ABB RobotStudio station: TPL2_Heredia_Biancuzzo.rspag

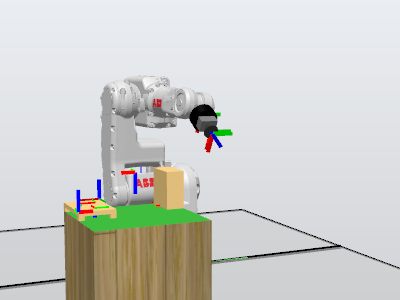
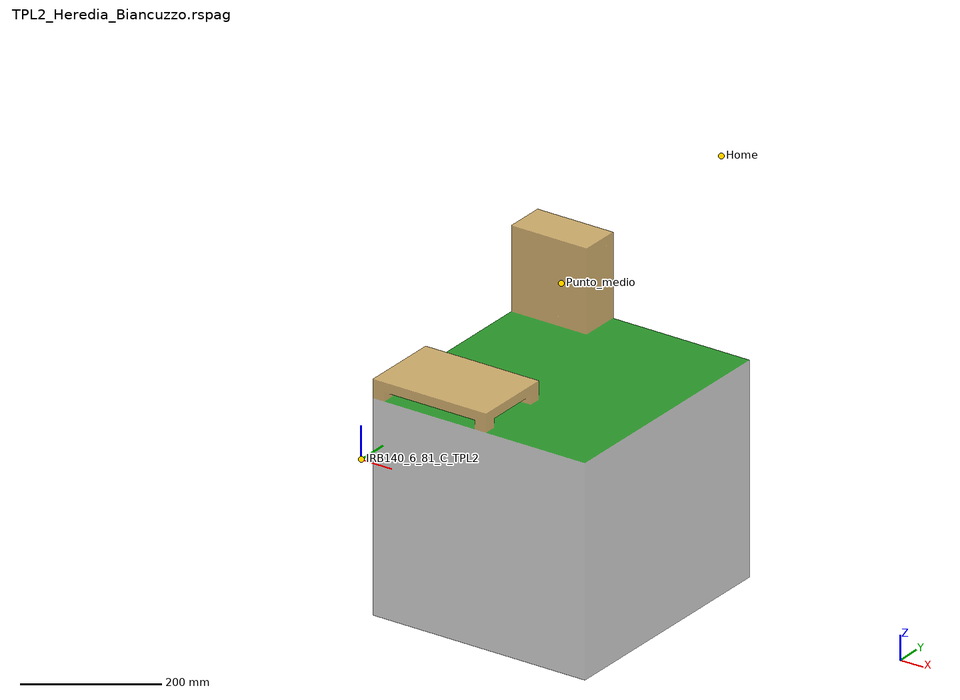
[picture v1: parts stored in the station drawn from their meshes, with robot base, taught points and paths (robot models come from the ABB library and are not in the file)]
--- station ---
Station Paletizado (saved by RobotStudio 25.5.11605.0)
Controller IRB140_6_81_TPL2
  mechanical unit ROB_1: IRB140_6_81_C_TPL2, 6 joints, base frame (0, 0, 0) mm
Layout (positions relative to the parent item):
  - Mesa [part], size 365 x 405 x 340 mm
  - Pallet [part], size 195 x 130 x 30 mm
  - Pieza1 [part], size 130 x 65 x 15 mm
  - Pieza2 [part], size 130 x 65 x 15 mm
  - Pieza3 [part], size 130 x 65 x 15 mm
  - Pieza4 [part], size 130 x 65 x 15 mm
  - Pieza5 [part], size 130 x 65 x 15 mm
  - Pieza6 [part], size 130 x 65 x 15 mm
  - Pieza7 [part], size 130 x 65 x 15 mm
  - Pieza8 [part], size 130 x 65 x 15 mm
  - Pieza9 [part], size 130 x 65 x 15 mm
  - Sopapa [mechanism] at (506.29, 39.79, 679.5) mm, rotated rx 180 ry 60 rz 180 deg
      TCP Sopapa at (0, -5, 103) mm
      links: Sopapa
  - IRB140_6_81_C_TPL2 [mechanism, from %ABB.RobotStudio.Models.IRB140%\IRB140_6_81_C_G_03.rslib] at (0, 0, 0) mm; joint values [0.0882, 0.0049, -0.0049, -0.1514, 0.5303, 0.175] (rad or m)
Attachment: Sopapa is attached to IRB140_6_81_C_TPL2 / Link6
Collision set Conjunto de colisión_1: Pieza1, Pieza2, Pieza3, Pieza4, Pieza5, Pieza6, Pieza7, Pieza8, Pieza9, Pallet, Mesa against IRB140_6_81_C_TPL2, Sopapa, near miss 0 m
EventTableEntry 2577: Group=, Trigger=DO_Sopapa 2578, Actions=[EventTableActionAttach 2579], Comment=, ActivationMode=2, Cyclic=false
EventTableTriggerIO 2578: IOValue=[1], IRC5Controller=? -1, Operator=0, SignalSource=IRB140_6_81_TPL2 1258
EventTableActionAttach 2579: AttachmentParent=Sopapa 1252, AttachmentChild=? -1, MountObject=false, Offset=[X=1, Y=0, Z=0, W=0, X=0, Y=1, Z=0, W=0, X=0, Y=0, Z=1, W=0, X=0, Y=0, Z=0, W=1], FlangeIndext=0, FindNearest=true
EventTableEntry 2580: Group=, Trigger=DO_Sopapa 2581, Actions=[EventTableActionDetach 2582], Comment=, ActivationMode=2, Cyclic=false
EventTableTriggerIO 2581: IOValue=[0], IRC5Controller=? -1, Operator=0, SignalSource=IRB140_6_81_TPL2 1258
EventTableActionDetach 2582: AttachmentParent=Sopapa 1252, AttachmentChild=? -1

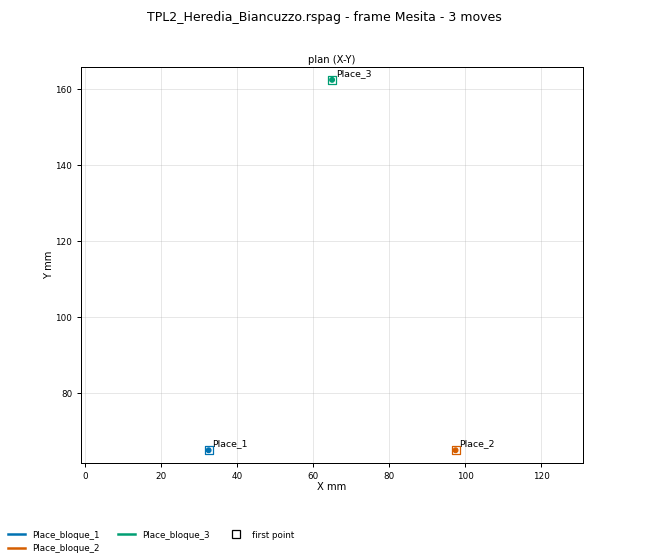
[picture p0: tool path of TPL2_Heredia_Biancuzzo.rspag in frame Mesita, 3 of 18 moves have a stored position in this frame; points joined in program order, loops and branches not executed]
--- Backups/IRB140_6_81_TPL2/RAPID/TASK1/PROGMOD/CalibData.mod ---
MODULE CalibData

ENDMODULE

--- Backups/IRB140_6_81_TPL2/RAPID/TASK1/PROGMOD/Module1.mod ---
MODULE Module1
    PERS wobjdata Mesa:=[FALSE,TRUE,"",[[300,5,340],[0.707107,0,0,-0.707107]],[[0,0,0],[1,0,0,0]]];
    PERS wobjdata Mesita:=[FALSE,TRUE,"",[[300,-270,370],[0.707107,0,0,-0.707107]],[[0,0,30],[1,0,0,0]]];

    PERS tooldata Sopapa:=[TRUE,[[0,-5,103],[1,0,0,0]],[0.5,[0,0,40],[1,0,0,0],0,0,0]];
    PERS tooldata SopapaBloque:=[TRUE,[[0,-5,118],[1,0,0,0]],[0.5,[0,0,40],[1,0,0,0],0,0,0]];

    CONST robtarget Mesita_og:=[[275,0,30],[1,0,0,0],[0,0,0,0],[9E+09,9E+09,9E+09,9E+09,9E+09,9E+09]];
    CONST robtarget Mesita_impar:=[[130,195,0],[0,0,0,1],[0,0,0,0],[9E+09,9E+09,9E+09,9E+09,9E+09,9E+09]];
    CONST robtarget Mesita_par:=[[0,0,0],[1,0,0,0],[0,0,0,0],[9E+09,9E+09,9E+09,9E+09,9E+09,9E+09]];

    CONST robtarget Home:=[[595.492,34.789,628],[0.5,0,0.866025404,0],[0,0,0,0],[9E+09,9E+09,9E+09,9E+09,9E+09,9E+09]];
    CONST robtarget Punto_medio:=[[482.5,-197.5,490],[0,-0.707106781,0.707106781,0],[0,0,0,0],[9E+09,9E+09,9E+09,9E+09,9E+09,9E+09]];

    CONST robtarget Pick_base:=[[32.5,65,0],[0,1,0,0],[0,0,0,0],[9E+09,9E+09,9E+09,9E+09,9E+09,9E+09]];
    CONST robtarget Place_1:=[[32.5,65,0],[0,1,0,0],[0,0,0,0],[9E+09,9E+09,9E+09,9E+09,9E+09,9E+09]];
    CONST robtarget Place_2:=[[97.5,65,0],[0,0,1,0],[0,0,0,0],[9E+09,9E+09,9E+09,9E+09,9E+09,9E+09]];
    CONST robtarget Place_3:=[[65,162.5,0],[0,-0.707106781,0.707106781,0],[0,0,0,0],[9E+09,9E+09,9E+09,9E+09,9E+09,9E+09]];

    CONST intnum Offset_soltar := 0;
    CONST intnum Offset_pick := 40;
    CONST intnum Offset_place := 40;
    CONST intnum Offset_diag := 10;

    CONST intnum Altura_bloque := 15;

    VAR intnum Cajas_en_pallet := 0;
    VAR intnum Cant_pallet := 9;
    VAR intnum Cant_bloques := 9;

    PROC main()

        Mesita.uframe := PoseMult(Mesa.uframe, [Mesita_og.trans, Mesita_og.rot]);
        SopapaBloque.tframe := PoseMult(Sopapa.tframe, [[0, 0, Altura_bloque + Offset_soltar], [1, 0, 0, 0]]);

        ! TPErase;
        ! TPReadNum Cajas_en_pallet, "¿Cuantas cajas hay en el pallet?";

        Cajas_en_pallet := 2;

        MoveJ Home,v100,z100,Sopapa\WObj:=wobj0;
        Desactivar_sopapa;

        TPL2;

        MoveJ Home,v100,fine,Sopapa\WObj:=wobj0;
        Desactivar_sopapa;
    ENDPROC

    PROC TPL2()
        VAR intnum Contador_bloque;
        VAR intnum Nivel;
        VAR robtarget Oframe;

        FOR i FROM Cajas_en_pallet TO Min(Cant_bloques, Cant_pallet) - 1 DO
            Pick_bloque Cant_bloques - i;
            Nivel := Trunc(i / 3);

            IF Nivel MOD 2 = 0 THEN
                Oframe := Offs(Mesita_par, 0, 0, Nivel * Altura_bloque);
            ELSE
                Oframe := Offs(Mesita_impar, 0, 0, Nivel * Altura_bloque);
            ENDIF
            Mesita.oframe := [Oframe.trans, Oframe.rot];

            ! Punto intermedio para evitar una colision con los bloques
            MoveJ Punto_medio,v100,z100,Sopapa\WObj:=wobj0;

            Contador_bloque := i MOD 3;
            IF Contador_bloque = 0 THEN
                Place_bloque_1;
            ELSEIF Contador_bloque = 1 THEN
                Place_bloque_2;
            ELSE
                Place_bloque_3;
            ENDIF

            MoveJ Punto_medio,v100,fine,Sopapa\WObj:=wobj0;
        ENDFOR

    ENDPROC

    PROC Pick_bloque(intnum Cant_stack)
        VAR intnum Offset_bloque;

        Offset_bloque := Cant_stack * Altura_bloque;
        MoveJ Offs(Pick_base, 0, 0, Offset_bloque + Offset_pick),v200,z100,Sopapa\WObj:=Mesa;
        MoveL Offs(Pick_base, 0, 0, Offset_bloque),v100,fine,Sopapa\WObj:=Mesa;
        Activar_sopapa;
        MoveL Offs(Pick_base, 0, 0, Offset_bloque + Offset_pick),v100,z100,Sopapa\WObj:=Mesa;
    ENDPROC

    PROC Place_bloque_1()
        MoveJ Offs(Place_1, 0, 0, Offset_place),v200,z100,SopapaBloque\WObj:=Mesita;
        MoveL Place_1,v100,fine,SopapaBloque\WObj:=Mesita;
        Desactivar_sopapa;
        MoveL Offs(Place_1, 0, 0, Offset_place),v100,z100,SopapaBloque\WObj:=Mesita;
    ENDPROC

    PROC Place_bloque_2()
        MoveJ Offs(Place_2, Offset_diag, 0, Offset_place),v200,z100,SopapaBloque\WObj:=Mesita;
        MoveL Offs(Place_2, Offset_diag, 0, Offset_diag),v100,z10,SopapaBloque\WObj:=Mesita;
        MoveL Place_2,v100,fine,SopapaBloque\WObj:=Mesita;
        Desactivar_sopapa;
        MoveL Offs(Place_2, 0, 0, Offset_place),v100,z100,SopapaBloque\WObj:=Mesita;
    ENDPROC

    PROC Place_bloque_3()
        MoveJ Offs(Place_3, 0, Offset_diag, Offset_place),v200,z100,SopapaBloque\WObj:=Mesita;
        MoveL Offs(Place_3, 0, Offset_diag, Offset_diag),v100,z10,SopapaBloque\WObj:=Mesita;
        MoveL Place_3,v100,fine,SopapaBloque\WObj:=Mesita;
        Desactivar_sopapa;
        MoveL Offs(Place_3, 0, 0, Offset_place),v100,z100,SopapaBloque\WObj:=Mesita;
    ENDPROC

    PROC Activar_sopapa()
        SetDO DO_Sopapa, 1;
        WaitTime 1;
    ENDPROC
    PROC Desactivar_sopapa()
        SetDO DO_Sopapa, 0;
        WaitTime 1;
    ENDPROC
ENDMODULE

--- Backups/IRB140_6_81_TPL2/SYSPAR/EIO.cfg ---
EIO:CFG_1.0:6:1::
#
EIO_SIGNAL:

      -Name "DO_Sopapa" -SignalType "DO"
